Fanuc TP program (LS listing): ManyMo.LS

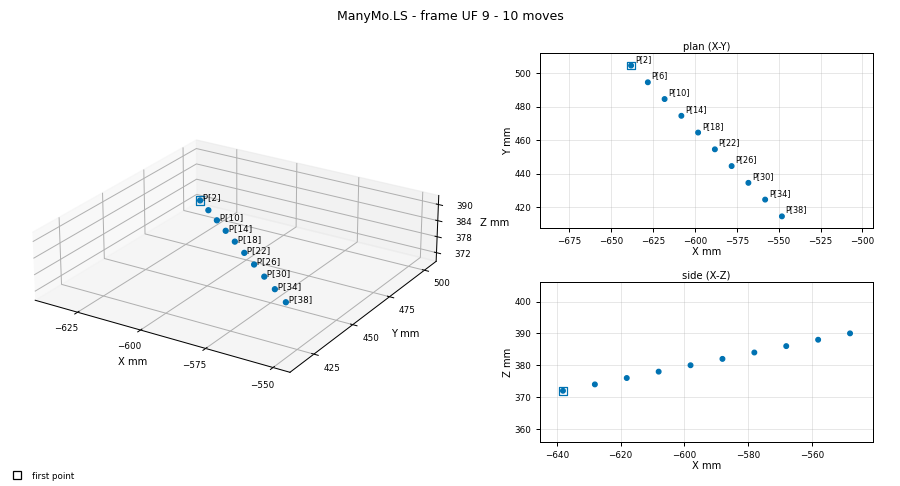
[picture p0: tool path of ManyMo.LS in frame UF 9, 10 of 40 moves have a stored position in this frame; points joined in program order, loops and branches not executed]
/PROG  ManyMo
/ATTR
OWNER		= MNEDITOR;
COMMENT		= "RoboDK sequence";
PROG_SIZE	= 0;
CREATE		= DATE 31-12-14  TIME 12:00:00;
MODIFIED	= DATE 31-12-14  TIME 12:00:00;
FILE_NAME	= ManyMo;
VERSION		= 0;
LINE_COUNT	= 59;
MEMORY_SIZE	= 0;
PROTECT		= READ_WRITE;
TCD:  STACK_SIZE	= 0,
      TASK_PRIORITY	= 50,
      TIME_SLICE	= 0,
      BUSY_LAMP_OFF	= 0,
      ABORT_REQUEST	= 0,
      PAUSE_REQUEST	= 0;
DEFAULT_GROUP	= 1,*,*,*,*;
CONTROL_CODE	= 00000000 00000000;
/MN
   1:  ! Program generated by RoboDK v6.0.7 for Fanuc M-1iA/0.5S on XX ;
   2:  ! /XX/XXXX 18:00:00 ;
   3:  ! Using nominal kinematics. ;
   4:  PR[9,1]=1234.570 ;
   5:  PR[9,2]=-98.765 ;
   6:  PR[9,3]=50.500 ;
   7:  PR[9,4]=0.000 ;
   8:  PR[9,5]=0.000 ;
   9:  PR[9,6]=30.000 ;
  10:  UFRAME[9]=PR[9] ;
  11:  UFRAME_NUM=9 ;
  12:  PR[9,1]=10.000 ;
  13:  PR[9,2]=20.000 ;
  14:  PR[9,3]=150.000 ;
  15:  PR[9,4]=0.000 ;
  16:  PR[9,5]=0.000 ;
  17:  PR[9,6]=0.000 ;
  18:  UTOOL[9]=PR[9] ;
  19:  UTOOL_NUM=9 ;
  20:J P[1] 10% FINE ;
  21:L P[2] 500mm/sec FINE ;
  22:J P[3] 10% FINE ;
  23:L P[4] 500mm/sec FINE ;
  24:J P[5] 10% FINE ;
  25:L P[6] 500mm/sec FINE ;
  26:J P[7] 10% FINE ;
  27:L P[8] 500mm/sec FINE ;
  28:J P[9] 10% FINE ;
  29:L P[10] 500mm/sec FINE ;
  30:J P[11] 10% FINE ;
  31:L P[12] 500mm/sec FINE ;
  32:J P[13] 10% FINE ;
  33:L P[14] 500mm/sec FINE ;
  34:J P[15] 10% FINE ;
  35:L P[16] 500mm/sec FINE ;
  36:J P[17] 10% FINE ;
  37:L P[18] 500mm/sec FINE ;
  38:J P[19] 10% FINE ;
  39:L P[20] 500mm/sec FINE ;
  40:J P[21] 10% FINE ;
  41:L P[22] 500mm/sec FINE ;
  42:J P[23] 10% FINE ;
  43:L P[24] 500mm/sec FINE ;
  44:J P[25] 10% FINE ;
  45:L P[26] 500mm/sec FINE ;
  46:J P[27] 10% FINE ;
  47:L P[28] 500mm/sec FINE ;
  48:J P[29] 10% FINE ;
  49:L P[30] 500mm/sec FINE ;
  50:J P[31] 10% FINE ;
  51:L P[32] 500mm/sec FINE ;
  52:J P[33] 10% FINE ;
  53:L P[34] 500mm/sec FINE ;
  54:J P[35] 10% FINE ;
  55:L P[36] 500mm/sec FINE ;
  56:J P[37] 10% FINE ;
  57:L P[38] 500mm/sec FINE ;
  58:J P[39] 10% FINE ;
  59:L P[40] 500mm/sec FINE ;
/POS
P[1]{
   GP1:
    UF : 9, UT : 9,
	J1=    10.000000 deg,	J2=    -20.000000 deg,	J3=    50.000000  mm,
	J4=    30.000000 deg
};
P[2]{
   GP1:
    UF : 9, UT : 9,        CONFIG : 'L, 0, 0, 0',
	X =  -638.084  mm,	Y =   504.480  mm,	Z =   372.034  mm,
	W =  -165.000 deg,	P =    50.000 deg,	R =   150.000 deg
};
P[3]{
   GP1:
    UF : 9, UT : 9,
	J1=    30.000000 deg,	J2=    25.000000 deg,	J3=    80.000000  mm,
	J4=    -45.000000 deg
};
P[4]{
   GP1:
    UF : 9, UT : 9,
	J1=    10.000000 deg,	J2=    -20.000000 deg,	J3=    50.000000  mm,
	J4=    30.000000 deg
};
P[5]{
   GP1:
    UF : 9, UT : 9,
	J1=    10.000000 deg,	J2=    -20.000000 deg,	J3=    50.000000  mm,
	J4=    30.000000 deg
};
P[6]{
   GP1:
    UF : 9, UT : 9,        CONFIG : 'L, 0, 0, 0',
	X =  -628.084  mm,	Y =   494.480  mm,	Z =   374.034  mm,
	W =  -165.000 deg,	P =    50.000 deg,	R =   150.000 deg
};
P[7]{
   GP1:
    UF : 9, UT : 9,
	J1=    30.000000 deg,	J2=    25.000000 deg,	J3=    80.000000  mm,
	J4=    -45.000000 deg
};
P[8]{
   GP1:
    UF : 9, UT : 9,
	J1=    10.000000 deg,	J2=    -20.000000 deg,	J3=    50.000000  mm,
	J4=    30.000000 deg
};
P[9]{
   GP1:
    UF : 9, UT : 9,
	J1=    10.000000 deg,	J2=    -20.000000 deg,	J3=    50.000000  mm,
	J4=    30.000000 deg
};
P[10]{
   GP1:
    UF : 9, UT : 9,        CONFIG : 'L, 0, 0, 0',
	X =  -618.084  mm,	Y =   484.480  mm,	Z =   376.034  mm,
	W =  -165.000 deg,	P =    50.000 deg,	R =   150.000 deg
};
P[11]{
   GP1:
    UF : 9, UT : 9,
	J1=    30.000000 deg,	J2=    25.000000 deg,	J3=    80.000000  mm,
	J4=    -45.000000 deg
};
P[12]{
   GP1:
    UF : 9, UT : 9,
	J1=    10.000000 deg,	J2=    -20.000000 deg,	J3=    50.000000  mm,
	J4=    30.000000 deg
};
P[13]{
   GP1:
    UF : 9, UT : 9,
	J1=    10.000000 deg,	J2=    -20.000000 deg,	J3=    50.000000  mm,
	J4=    30.000000 deg
};
P[14]{
   GP1:
    UF : 9, UT : 9,        CONFIG : 'L, 0, 0, 0',
	X =  -608.084  mm,	Y =   474.480  mm,	Z =   378.034  mm,
	W =  -165.000 deg,	P =    50.000 deg,	R =   150.000 deg
};
P[15]{
   GP1:
    UF : 9, UT : 9,
	J1=    30.000000 deg,	J2=    25.000000 deg,	J3=    80.000000  mm,
	J4=    -45.000000 deg
};
P[16]{
   GP1:
    UF : 9, UT : 9,
	J1=    10.000000 deg,	J2=    -20.000000 deg,	J3=    50.000000  mm,
	J4=    30.000000 deg
};
P[17]{
   GP1:
    UF : 9, UT : 9,
	J1=    10.000000 deg,	J2=    -20.000000 deg,	J3=    50.000000  mm,
	J4=    30.000000 deg
};
P[18]{
   GP1:
    UF : 9, UT : 9,        CONFIG : 'L, 0, 0, 0',
	X =  -598.084  mm,	Y =   464.480  mm,	Z =   380.034  mm,
	W =  -165.000 deg,	P =    50.000 deg,	R =   150.000 deg
};
P[19]{
   GP1:
    UF : 9, UT : 9,
	J1=    30.000000 deg,	J2=    25.000000 deg,	J3=    80.000000  mm,
	J4=    -45.000000 deg
};
P[20]{
   GP1:
    UF : 9, UT : 9,
	J1=    10.000000 deg,	J2=    -20.000000 deg,	J3=    50.000000  mm,
	J4=    30.000000 deg
};
P[21]{
   GP1:
    UF : 9, UT : 9,
	J1=    10.000000 deg,	J2=    -20.000000 deg,	J3=    50.000000  mm,
	J4=    30.000000 deg
};
P[22]{
   GP1:
    UF : 9, UT : 9,        CONFIG : 'L, 0, 0, 0',
	X =  -588.084  mm,	Y =   454.480  mm,	Z =   382.034  mm,
	W =  -165.000 deg,	P =    50.000 deg,	R =   150.000 deg
};
P[23]{
   GP1:
    UF : 9, UT : 9,
	J1=    30.000000 deg,	J2=    25.000000 deg,	J3=    80.000000  mm,
	J4=    -45.000000 deg
};
P[24]{
   GP1:
    UF : 9, UT : 9,
	J1=    10.000000 deg,	J2=    -20.000000 deg,	J3=    50.000000  mm,
	J4=    30.000000 deg
};
P[25]{
   GP1:
    UF : 9, UT : 9,
	J1=    10.000000 deg,	J2=    -20.000000 deg,	J3=    50.000000  mm,
	J4=    30.000000 deg
};
P[26]{
   GP1:
    UF : 9, UT : 9,        CONFIG : 'L, 0, 0, 0',
	X =  -578.084  mm,	Y =   444.480  mm,	Z =   384.034  mm,
	W =  -165.000 deg,	P =    50.000 deg,	R =   150.000 deg
};
P[27]{
   GP1:
    UF : 9, UT : 9,
	J1=    30.000000 deg,	J2=    25.000000 deg,	J3=    80.000000  mm,
	J4=    -45.000000 deg
};
P[28]{
   GP1:
    UF : 9, UT : 9,
	J1=    10.000000 deg,	J2=    -20.000000 deg,	J3=    50.000000  mm,
	J4=    30.000000 deg
};
P[29]{
   GP1:
    UF : 9, UT : 9,
	J1=    10.000000 deg,	J2=    -20.000000 deg,	J3=    50.000000  mm,
	J4=    30.000000 deg
};
P[30]{
   GP1:
    UF : 9, UT : 9,        CONFIG : 'L, 0, 0, 0',
	X =  -568.084  mm,	Y =   434.480  mm,	Z =   386.034  mm,
	W =  -165.000 deg,	P =    50.000 deg,	R =   150.000 deg
};
P[31]{
   GP1:
    UF : 9, UT : 9,
	J1=    30.000000 deg,	J2=    25.000000 deg,	J3=    80.000000  mm,
	J4=    -45.000000 deg
};
P[32]{
   GP1:
    UF : 9, UT : 9,
	J1=    10.000000 deg,	J2=    -20.000000 deg,	J3=    50.000000  mm,
	J4=    30.000000 deg
};
P[33]{
   GP1:
    UF : 9, UT : 9,
	J1=    10.000000 deg,	J2=    -20.000000 deg,	J3=    50.000000  mm,
	J4=    30.000000 deg
};
P[34]{
   GP1:
    UF : 9, UT : 9,        CONFIG : 'L, 0, 0, 0',
	X =  -558.084  mm,	Y =   424.480  mm,	Z =   388.034  mm,
	W =  -165.000 deg,	P =    50.000 deg,	R =   150.000 deg
};
P[35]{
   GP1:
    UF : 9, UT : 9,
	J1=    30.000000 deg,	J2=    25.000000 deg,	J3=    80.000000  mm,
	J4=    -45.000000 deg
};
P[36]{
   GP1:
    UF : 9, UT : 9,
	J1=    10.000000 deg,	J2=    -20.000000 deg,	J3=    50.000000  mm,
	J4=    30.000000 deg
};
P[37]{
   GP1:
    UF : 9, UT : 9,
	J1=    10.000000 deg,	J2=    -20.000000 deg,	J3=    50.000000  mm,
	J4=    30.000000 deg
};
P[38]{
   GP1:
    UF : 9, UT : 9,        CONFIG : 'L, 0, 0, 0',
	X =  -548.084  mm,	Y =   414.480  mm,	Z =   390.034  mm,
	W =  -165.000 deg,	P =    50.000 deg,	R =   150.000 deg
};
P[39]{
   GP1:
    UF : 9, UT : 9,
	J1=    30.000000 deg,	J2=    25.000000 deg,	J3=    80.000000  mm,
	J4=    -45.000000 deg
};
P[40]{
   GP1:
    UF : 9, UT : 9,
	J1=    10.000000 deg,	J2=    -20.000000 deg,	J3=    50.000000  mm,
	J4=    30.000000 deg
};
/END
